(* IEC 61131-3 sources: plc-st-test/test/security/fixtures/plugins/Tests, 1 file *)

(* ---- TEST_Never.st ---- *)
FUNCTION_BLOCK TEST_Never
VAR
  uut : FB_Dummy;
END_VAR
METHOD Test_NeverRuns
  ASSERT_EQUAL_DINT(uut.nValue, 0);
END_METHOD
END_FUNCTION_BLOCK
